(* IEC 61131-3 sources: LASAL/Network/TcpServer, 1 file *)

(* ---- ONE_TcpServer_Table.st ---- *)
#define OBJECTS_CONFIG

//Define part of class _TCPIP_SERVER
#ifndef OS_VERSION_MIN_SALAMANDER
    #define OS_VERSION_MIN_SALAMANDER          0x9000
  #endif
  #define TCP_SVR_NO_ERROR                          0

  #define TCP_SVR_ERR_INVALID_SOCKET            -1

  #define TCP_SVR_ERR_SET_PARA_INVALID_CMD     -10
  #define TCP_SVR_ERR_SET_PARA_INVALID_SUB_CMD -11

  #define TCP_SVR_ERR_TASK_ALREADY_EXIST       -12

  // - RETURN VALUES PRIVATE METHOD Read_AP_TaskPeriod
  #define TCP_SVR_ERR_TASK_TIME_NO_APP            -31
  #define TCP_SVR_ERR_TASK_TIME_WRONG_TASK_TYPE   -33
  #define TCP_SVR_ERR_TASK_TIME_OBJ_NOT_FOUND     -35

  // - RETURN VALUES PRIVATE METHOD Read_LSLOBJ_CRC32
  #define TCP_SVR_ERR_GET_LSLOBJ_NAME             -20
  #define TCP_SVR_ERR_INVALID_POINTER             -21

  // - RETURN VALUES PRIVATE METHOD AP_TaskCreate
  #define TCP_SVR_ERR_TASK_CREATE                 -40

  // - RETURN VALUES PRIVATE METHOD AP_SemaCreate
  #define TCP_SVR_ERR_SEMA_CREATE                 -50
  #define TCP_SVR_ERR_SEMA_INVALID_IDX            -51
  #define TCP_SVR_ERR_SEMA_INVALID_NAME           -52

  #define TCP_SVR_SEND_BUFFER_EMPTY               -6
  #define TCP_SVR_ERR_SEND_BUFFER_FATAL_ERROR     -7

  #define TCP_SVR_SEND_BUFFER_FULL      -4

  #define TCP_SVR_SOCK_INFO_CONNECT                 1
  #define TCP_SVR_SOCK_INFO_DISCONNECT              0

  #define TCP_SVR_ERR_GROUP_OS                      0
  #define TCP_SVR_ERR_GROUP_AP                      1

  #define TCP_SVR_ERR_CODE_AP_TIMEOUT              -1

  #ifndef INIT_FIRSTSCAN
    #define INIT_FIRSTSCAN                         12
  #endif

  #ifndef AP_TASK_PRIORITY_DEFAULT
    #define AP_TASK_PRIORITY_DEFAULT               14
  #endif

  #define TCP_SVR_ERR_MAIN_INIT                   -90

  #define TCP_SVR_ERR_MAX_CONN                    -80

  #ifndef KEEPALIVE_INTERVAL_DEFAULT
    #define KEEPALIVE_INTERVAL_DEFAULT           7200
  #endif

  #ifndef KEEPALIVE_RETRYTIME_DEFAULT
    #define KEEPALIVE_RETRYTIME_DEFAULT            75
  #endif

  #ifndef KEEPALIVE_RETRYCNT_DEFUALT
    #define KEEPALIVE_RETRYCNT_DEFUALT             10
  #endif

  #ifndef CLOSE_SOCKET_TYPE_DEFAULT
    #define CLOSE_SOCKET_TYPE_DEFAULT               0
  #endif
#include "..\..\Class\_TCPIP_SERVER\SalamanderDelay.h"
#include <.\lsl_st_mt.h>

FUNCTION GLOBAL TAB ONE_TcpServer
-1$UINT, 0$UINT,
0$UINT, 0$UINT,

8$UDINT,
TO_UDINT(916194998), "_CheckSum", 1$UINT, 0$UINT, 1$UINT,
TO_UDINT(26234884), "_TCPIP_SERVER", 1$UINT, 37$UINT, 0$UINT,
TO_UDINT(2047756655), "CommandRouter", 0$UINT, 0$UINT, 1$UINT,
TO_UDINT(1706127036), "CommandServer", 0$UINT, 0$UINT, 1$UINT,
TO_UDINT(2225119864), "MerkerEx", 1$UINT, 22$UINT, 3$UINT,
TO_UDINT(1850111279), "String", 1$UINT, 10$UINT, 3$UINT,
TO_UDINT(2898603620), "StringInternal", 1$UINT, 82$UINT, 0$UINT,
TO_UDINT(3232495061), "VirtualBaseInit", 1$UINT, 3$UINT, 0$UINT,

1$UINT, TO_UDINT(554147771), "COMMANDSERVER\_BASE\CHECKSUM",

_NO_ATTR, TO_UDINT(2047756655), "COMMANDROUTER",

_NO_ATTR, TO_UDINT(1706127036), "COMMANDSERVER",

1$UINT, TO_UDINT(2432255397), "COMMANDSERVER\_BASE\STRSEMANAME01\MERKEREX0",
1$UINT, TO_UDINT(152773540), "COMMANDSERVER\_BASE\STRSEMANAME02\MERKEREX0",
1$UINT, TO_UDINT(1469116870), "COMMANDSERVER\_BASE\STRTASKNAME\MERKEREX0",

1$UINT, TO_UDINT(2422395016), "COMMANDSERVER\_BASE\STRSEMANAME01",
1$UINT, TO_UDINT(158040370), "COMMANDSERVER\_BASE\STRSEMANAME02",
1$UINT, TO_UDINT(677430128), "COMMANDSERVER\_BASE\STRTASKNAME",

//Internal connections
0$UDINT,
7$UDINT,
TO_UDINT(2), "CheckSum", TO_UDINT(0),
TO_UDINT(2), "StrTaskName", TO_UDINT(8),
TO_UDINT(2), "StrSemaName01", TO_UDINT(6),
TO_UDINT(2), "StrSemaName02", TO_UDINT(7),
TO_UDINT(6), "MerkerEx0", TO_UDINT(3),
TO_UDINT(7), "MerkerEx0", TO_UDINT(4),
TO_UDINT(8), "MerkerEx0", TO_UDINT(5),
0$UDINT,
4$UDINT,
TO_UDINT(2), "CmdRouter", TO_UDINT(1), "CmdRouter",
TO_UDINT(6), "DataBuffer", TO_UDINT(3), "m_udLength",
TO_UDINT(7), "DataBuffer", TO_UDINT(4), "m_udLength",
TO_UDINT(8), "DataBuffer", TO_UDINT(5), "m_udLength",

//Initialization values
0$UDINT,
14$UDINT,
TO_UDINT(1), "Speed", TO_UDINT(10000000),//|TcpServer.commandRouter.Speed;
TO_UDINT(1), "Acc", TO_UDINT(40000000),//|TcpServer.commandRouter.Acc;
TO_UDINT(1), "YSpeed", TO_UDINT(50000000),//|TcpServer.commandRouter.YSpeed;
TO_UDINT(1), "YAcc", TO_UDINT(600000000),//|TcpServer.commandRouter.YAcc;
TO_UDINT(1), "Controller", TO_UDINT(MoveController::_Idle),//|TcpServer.commandRouter.Controller;
TO_UDINT(1), "clib", TO_UDINT(0),//|TcpServer.commandRouter.clib;
TO_UDINT(2), "cPort", TO_UDINT(1985),//|TcpServer.commandServer.cPort;
TO_UDINT(2), "cMaxConnections", TO_UDINT(0),//|TcpServer.commandServer.cMaxConnections;
TO_UDINT(3), "ThreadSafe", TO_UDINT(0),//|TcpServer.StrSemaName01\_base\commandServer\MerkerEx0.ThreadSafe;
TO_UDINT(4), "ThreadSafe", TO_UDINT(0),//|TcpServer.StrSemaName02\_base\commandServer\MerkerEx0.ThreadSafe;
TO_UDINT(5), "ThreadSafe", TO_UDINT(0),//|TcpServer.StrTaskName\_base\commandServer\MerkerEx0.ThreadSafe;
TO_UDINT(6), "SingleRealloc", TO_UDINT(1),//|TcpServer._base\commandServer\StrSemaName01.SingleRealloc;
TO_UDINT(7), "SingleRealloc", TO_UDINT(1),//|TcpServer._base\commandServer\StrSemaName02.SingleRealloc;
TO_UDINT(8), "SingleRealloc", TO_UDINT(1),//|TcpServer._base\commandServer\StrTaskName.SingleRealloc;

//Symbolic initialization values
0$UDINT,
0$UDINT,

//Initialization of string values
0$UDINT,
0$UDINT,

//Configuration of tasks (RealTime, Cyclic, Background)
0$UDINT,
0$UDINT,

0$UDINT,
1$UDINT,
TO_UDINT(2), (10)$UDINT, 4194303$DINT, 	//COMMANDSERVER

0$UDINT,
0$UDINT,

//External connections
0$UDINT,
1$UDINT,
TO_UDINT(1), "Controller", C_DIR, TO_UDINT(1841029985), "moveController","Status",

//Magic internal connections
0$UDINT,
0$UDINT,

//Configuration of timeslots of tasks (RealTime, Cyclic)
#ifdef __LSLLDR_TIMESLOTS__
0$UDINT,
0$UDINT,

0$UDINT,
0$UDINT,

#endif //__LSLLDR_TIMESLOTS__

//MultiMaster connections
#ifdef __LSLLDR_MULTIMASTER__
0$UDINT,
0$UDINT,
#endif //__LSLLDR_MULTIMASTER__

//Configuration for task ID (RealTime, CyclicTime)
#ifdef __LSLLDR_TASKID__
"\\\\TASKS2  "
0$UDINT,
0$UDINT,

0$UDINT,
1$UDINT,
(0)$UDINT, 	//COMMANDSERVER

0$UDINT,
0$UDINT,

#endif //__LSLLDR_TASKID__

END_FUNCTION
